{attribute 'qualified_only'}
VAR_GLOBAL
	
	_i_b_endSwitch_1 AT %I* :BOOL;
	_i_b_endSwitch_2 AT %I* :BOOL;
	_i_b_endSwitch_3 AT %I* :BOOL;
	_i_b_endSwitch_4 AT %I* :BOOL;
	_i_b_startButton AT %I*	:BOOL;
	_i_b_stopButton	 AT %I*	:BOOL;

	_o_b_valve1	AT %Q*	:BOOL;
	_o_b_valve2	AT %Q*	:BOOL;
	_o_b_valve3	AT %Q*	:BOOL;
	_o_b_valve4	AT %Q*	:BOOL;



END_VAR

(* stored: Version 1.1.0.1
   GVL IN_OUT: Id {9aa5e3e2-501b-4032-bbd8-190d0ac61ae1} *)
